Fanuc KAREL source: kt00741.KL

-- PROVISIONAL review KL for V770-1; original PC SHA256 8e042effa6b8be7742bac7b6c4b892eed9fd4109bc024c16455271a1cc0163e3
-- Incomplete behavior may be omitted. Consult companion uncertainty JSON. Do not deploy.
PROGRAM KT00741
%NOLOCKGROUP
VAR
  OUT : INTEGER
-- UNRESOLVED_DECL ARG type=002017
BEGIN
  -- UNRESOLVED_PC offsets 5-18; opcodes 22,1D,23
  -- UNRESOLVED_PC offsets 23-27; opcodes 7F
END KT00741
